(* Logix 5000 project; controller R400_500_XLS vendor 1 type 14 code 216 rev 31.11; software revision 31.01; part 28 of 32 *)
(* tags used below, declared in another part *)
   Abort1 : DINT;   // Not Used
   Ashutdown : SINT;   // Not Used
   CycExcBuffer : UDT_CYCLE;
   CycleSequence : UDT_CYCLE_SEQUENCE;
   CycleTime : DINT[11];   // Last cycle time saved in seconds
   DrnSmp : DINT;
   DRYING : DINT;   // Drying id number
   FC05_ONS : DINT;
   FINALRINSE_1 : DINT;   // Final rinse 1 id number
   FINALRINSE_9 : DINT;   // Final rinse 9 id number
   iDecimalSeparatorIndex : INT;
   M : DINT[5];   // Memory Bits
   New_Value : SINT;
   ONS_FC05 : DINT;
   ONS_FC64 : DINT;
   Print_Data : BOOL;   // Print Treatment data
   print_Door_opened_template : STRING;   // Template for the door opened message
   print_Header_template : STRING[6];   // Template for the cycle header
   Print_Speed_Water : BOOL;
   Print_TreatEnd_Start_Data : BOOL;   // 2nd treatment of the cycle is started, pirnt Treatment Completed and Treatment data
   Print_TreatStart_Data : BOOL;   // Cycle is started Print start time and treatment data of the first treatment of the cycle
   PrintBufferInjectionRate : REAL;
   printTreatString : STRING[85];   // Treatment String
   PWR_PrintBuffer : UDT_WASH;
   rBuffer : REAL[4];
   rIn_WSH61 : REAL;
   Run : DINT;
   sCRLF : STRING;
   sDecimalSeparator : STRING;
   sFll_Zero : STRING[20];
   sOut_WSH61 : STRING;
   sPrntArray : STRING[300];   // Printer String Array
   SRE3_Serial_Number : STRING;   // Serial number
   String : STRING[50];   // String
   String_Temp : STRING;
   Tmr : TIMER[107];
   Trt_PrWsh : DINT;
   WASH_1 : DINT;   // Wash 1 id number
   WASH_5 : DINT;   // Wash 5 id number
   WSH36_SecondsRemaining : DINT;
   WSH36_TotalMinutesRemaining : DINT;
   WSH36_TotalSecondsRemaining : DINT;
   WSH41_Door_opened : STRING;
   WSH41_End_signal : BOOL;   // End of cycle signal
   WSH41_Header : STRING[6];   // The header being transferred to the print queue.
   WSH41_Hour : DINT;
   WSH41_Minute : DINT;
   WSH41_ONS : SINT;
   WSH41_Second : DINT;
   WSH41_Start_signal : BOOL;   // Start cycle signal One shot rising edge
   WSH41_Temp_time : STRING[3];
   WSH41_Time_template : STRING;
   WSH41_Total_minute : DINT;
   WSH41_Total_second : DINT;
   WSH41_Total_time : STRING;
   WSH41_Zero : STRING;
   ChemConcUnit : BOOL;   // 0 = mL/L; 1 = oz/gal
   ChemicalName : STRING[9];   // Used by HMI
   CurrentUser : STRING;   // Current User
   CycleName : STRING[12];
   CyclePtr : DINT;   // Cycle Pointeur
   ENABLE : BOOL;   // Enable bit
   I_Ld_Dr_Cls_Sw : BOOL;   // Load door close
   I_Unld_Dr_Cls_Sw : BOOL;   // Unload door close
   MaintainOpenLd : BOOL;
   MaintainOpenUnld : BOOL;
   PrintIndex : DINT;
   RcvryWtrTemp : DINT;
   sCycleCounter : STRING;
   sDate : STRING;   // String current date
   sTime : STRING;   // String current time
   SumpTemp : REAL;   // Sump temperature in °C
   TempUnit : BOOL;   // Temperature Units 0= Celcius 1 = Farhenheit
   Unit : Hrdwre;   // Unit Configuration
   UnLoad : Doors;
(* MainProgram, continued *)

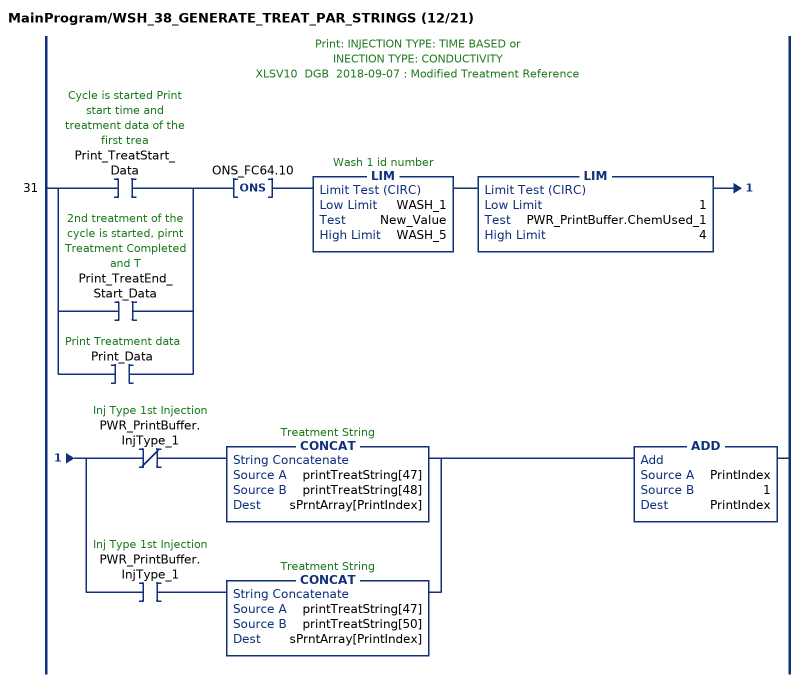
   [picture p570: MainProgram/WSH_38_GENERATE_TREAT_PAR_STRINGS rungs 31-31]
   // Print: INJECTION TYPE: TIME BASED or
   // INECTION TYPE: CONDUCTIVITY
   // XLSV10  DGB  2018-09-07 : Modified Treatment Reference
   31: [XIC(Print_TreatStart_Data) ,XIC(Print_TreatEnd_Start_Data) ,XIC(Print_Data) ]ONS(ONS_FC64.10)LIM(WASH_1,New_Value,WASH_5)LIM(1,PWR_PrintBuffer.ChemUsed_1,4)[XIO(PWR_PrintBuffer.InjType_1) CONCAT(printTreatString[47],printTreatString[48],sPrntArray[PrintIndex]) ,XIC(PWR_PrintBuffer.InjType_1) CONCAT(printTreatString[47],printTreatString[50],sPrntArray[PrintIndex]) ]ADD(PrintIndex,1,PrintIndex);
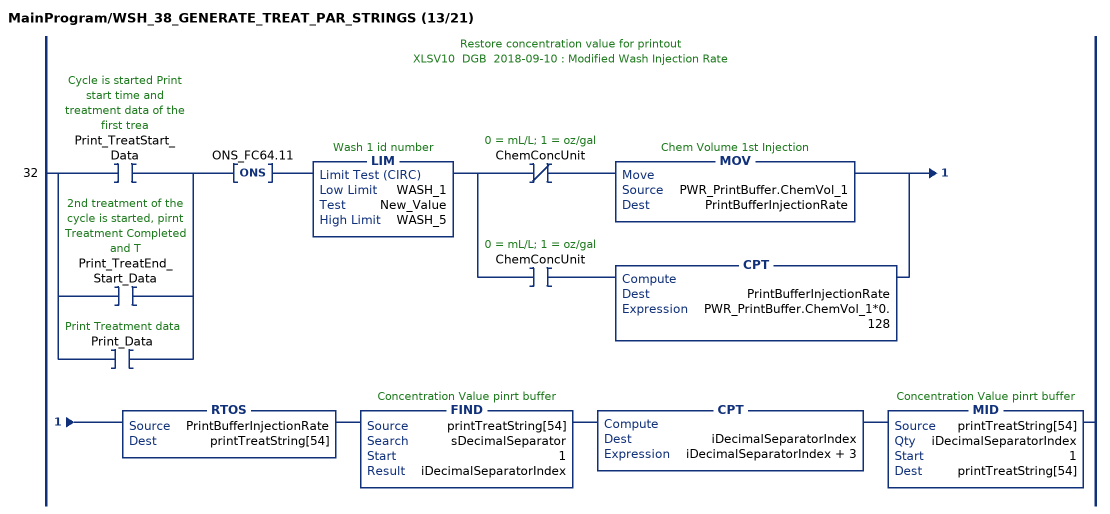
   // Restore concentration value for printout
   // XLSV10  DGB  2018-09-10 : Modified Wash Injection Rate
   32: [XIC(Print_TreatStart_Data) ,XIC(Print_TreatEnd_Start_Data) ,XIC(Print_Data) ]ONS(ONS_FC64.11)LIM(WASH_1,New_Value,WASH_5)[XIO(ChemConcUnit) MOV(PWR_PrintBuffer.ChemVol_1,PrintBufferInjectionRate) ,XIC(ChemConcUnit) CPT(PrintBufferInjectionRate,PWR_PrintBuffer.ChemVol_1*0.128) ]RTOS(PrintBufferInjectionRate,printTreatString[54])FIND(printTreatString[54],sDecimalSeparator,1,iDecimalSeparatorIndex)CPT(iDecimalSeparatorIndex,iDecimalSeparatorIndex + 3)MID(printTreatString[54],iDecimalSeparatorIndex,1,printTreatString[54]);
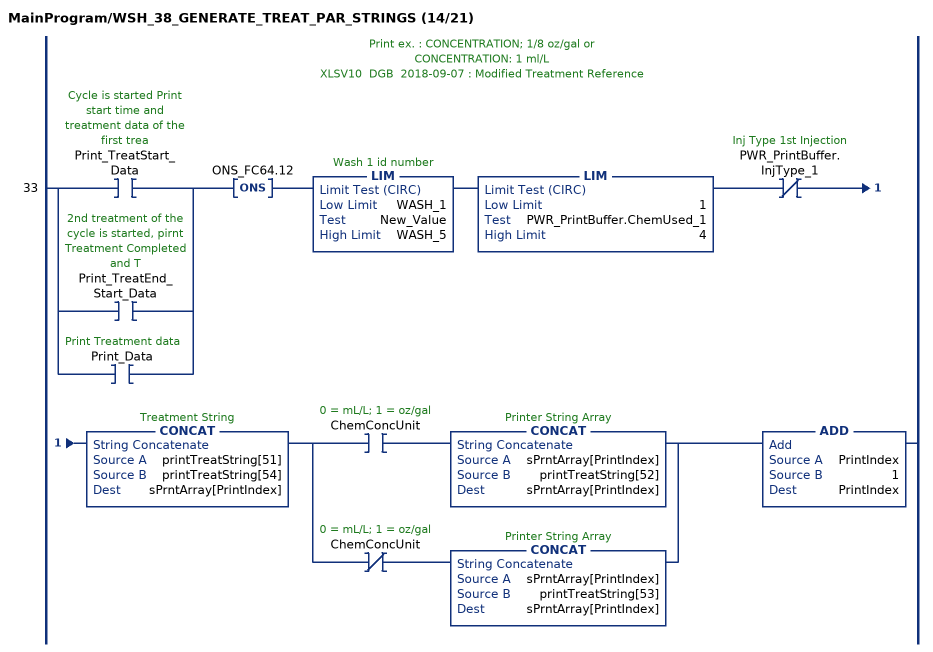
   // Print ex. : CONCENTRATION; 1/8 oz/gal or
   //         CONCENTRATION: 1 ml/L
   // XLSV10  DGB  2018-09-07 : Modified Treatment Reference
   33: [XIC(Print_TreatStart_Data) ,XIC(Print_TreatEnd_Start_Data) ,XIC(Print_Data) ]ONS(ONS_FC64.12)LIM(WASH_1,New_Value,WASH_5)LIM(1,PWR_PrintBuffer.ChemUsed_1,4)XIO(PWR_PrintBuffer.InjType_1)CONCAT(printTreatString[51],printTreatString[54],sPrntArray[PrintIndex])[XIC(ChemConcUnit) CONCAT(sPrntArray[PrintIndex],printTreatString[52],sPrntArray[PrintIndex]) ,XIO(ChemConcUnit) CONCAT(sPrntArray[PrintIndex],printTreatString[53],sPrntArray[PrintIndex]) ]ADD(PrintIndex,1,PrintIndex);
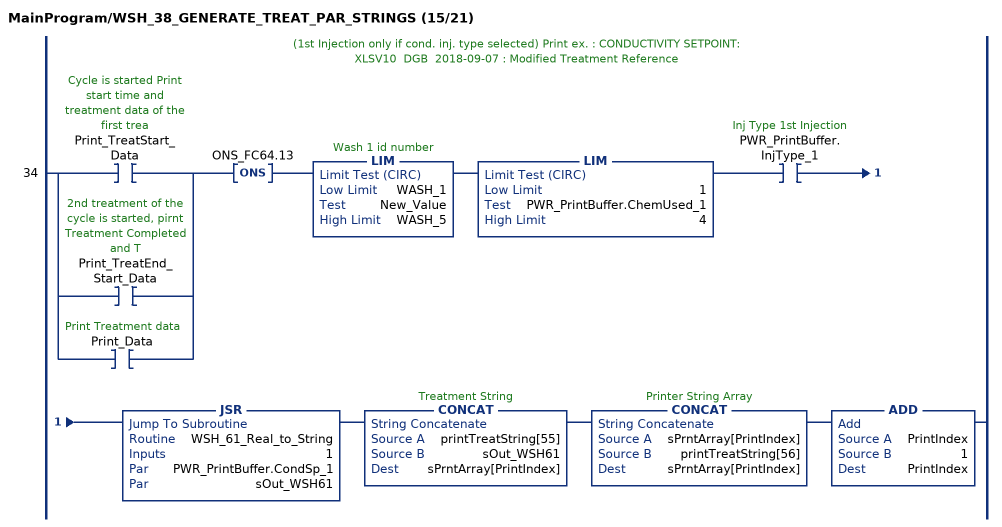
   // (1st Injection only if cond. inj. type selected) Print ex. : CONDUCTIVITY SETPOINT:
   // XLSV10  DGB  2018-09-07 : Modified Treatment Reference
   34: [XIC(Print_TreatStart_Data) ,XIC(Print_TreatEnd_Start_Data) ,XIC(Print_Data) ]ONS(ONS_FC64.13)LIM(WASH_1,New_Value,WASH_5)LIM(1,PWR_PrintBuffer.ChemUsed_1,4)XIC(PWR_PrintBuffer.InjType_1)JSR(WSH_61_Real_to_String,1,PWR_PrintBuffer.CondSp_1,sOut_WSH61)CONCAT(printTreatString[55],sOut_WSH61,sPrntArray[PrintIndex])CONCAT(sPrntArray[PrintIndex],printTreatString[56],sPrntArray[PrintIndex])ADD(PrintIndex,1,PrintIndex);
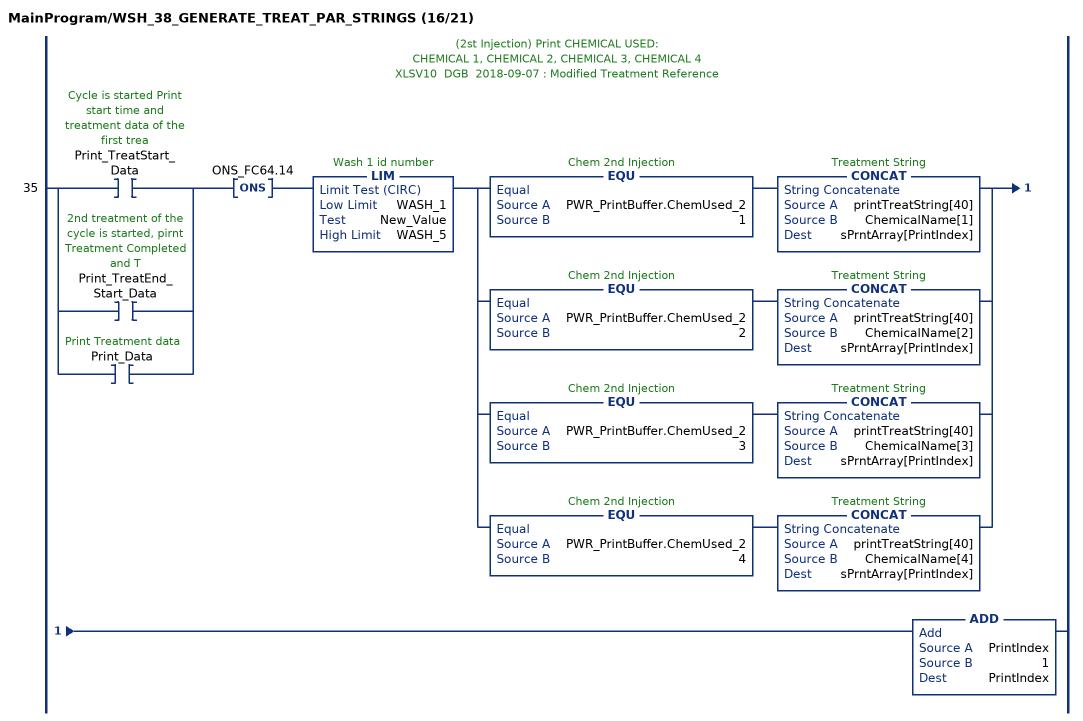
   // (2st Injection) Print CHEMICAL USED:
   //  CHEMICAL 1, CHEMICAL 2, CHEMICAL 3, CHEMICAL 4
   // XLSV10  DGB  2018-09-07 : Modified Treatment Reference
   35: [XIC(Print_TreatStart_Data) ,XIC(Print_TreatEnd_Start_Data) ,XIC(Print_Data) ]ONS(ONS_FC64.14)LIM(WASH_1,New_Value,WASH_5)[EQU(PWR_PrintBuffer.ChemUsed_2,1) CONCAT(printTreatString[40],ChemicalName[1],sPrntArray[PrintIndex]) ,EQU(PWR_PrintBuffer.ChemUsed_2,2) CONCAT(printTreatString[40],ChemicalName[2],sPrntArray[PrintIndex]) ,EQU(PWR_PrintBuffer.ChemUsed_2,3) CONCAT(printTreatString[40],ChemicalName[3],sPrntArray[PrintIndex]) ,EQU(PWR_PrintBuffer.ChemUsed_2,4) CONCAT(printTreatString[40],ChemicalName[4],sPrntArray[PrintIndex]) ]ADD(PrintIndex,1,PrintIndex);
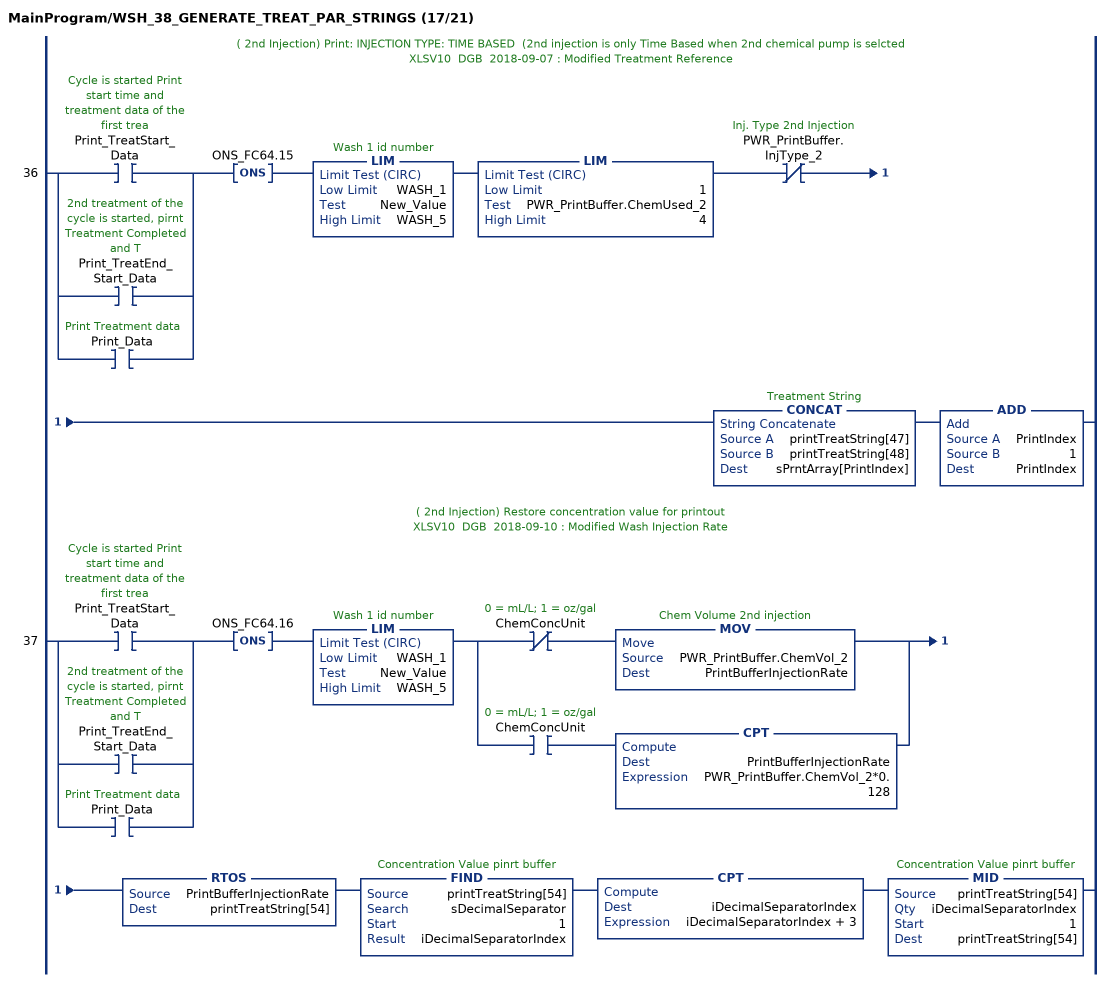
   // ( 2nd Injection) Print: INJECTION TYPE: TIME BASED  (2nd injection is only Time Based when 2nd chemical pump is selcted
   // XLSV10  DGB  2018-09-07 : Modified Treatment Reference
   36: [XIC(Print_TreatStart_Data) ,XIC(Print_TreatEnd_Start_Data) ,XIC(Print_Data) ]ONS(ONS_FC64.15)LIM(WASH_1,New_Value,WASH_5)LIM(1,PWR_PrintBuffer.ChemUsed_2,4)XIO(PWR_PrintBuffer.InjType_2)CONCAT(printTreatString[47],printTreatString[48],sPrntArray[PrintIndex])ADD(PrintIndex,1,PrintIndex);
   // ( 2nd Injection) Restore concentration value for printout
   // XLSV10  DGB  2018-09-10 : Modified Wash Injection Rate
   37: [XIC(Print_TreatStart_Data) ,XIC(Print_TreatEnd_Start_Data) ,XIC(Print_Data) ]ONS(ONS_FC64.16)LIM(WASH_1,New_Value,WASH_5)[XIO(ChemConcUnit) MOV(PWR_PrintBuffer.ChemVol_2,PrintBufferInjectionRate) ,XIC(ChemConcUnit) CPT(PrintBufferInjectionRate,PWR_PrintBuffer.ChemVol_2*0.128) ]RTOS(PrintBufferInjectionRate,printTreatString[54])FIND(printTreatString[54],sDecimalSeparator,1,iDecimalSeparatorIndex)CPT(iDecimalSeparatorIndex,iDecimalSeparatorIndex + 3)MID(printTreatString[54],iDecimalSeparatorIndex,1,printTreatString[54]);
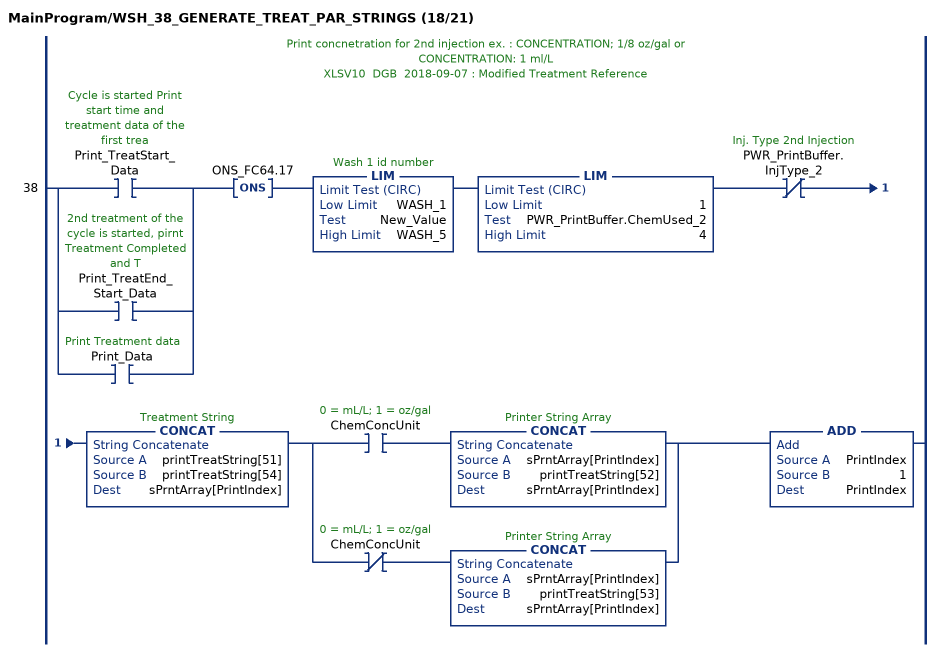
   // Print concnetration for 2nd injection ex. : CONCENTRATION; 1/8 oz/gal or
   //         CONCENTRATION: 1 ml/L
   // XLSV10  DGB  2018-09-07 : Modified Treatment Reference
   38: [XIC(Print_TreatStart_Data) ,XIC(Print_TreatEnd_Start_Data) ,XIC(Print_Data) ]ONS(ONS_FC64.17)LIM(WASH_1,New_Value,WASH_5)LIM(1,PWR_PrintBuffer.ChemUsed_2,4)XIO(PWR_PrintBuffer.InjType_2)CONCAT(printTreatString[51],printTreatString[54],sPrntArray[PrintIndex])[XIC(ChemConcUnit) CONCAT(sPrntArray[PrintIndex],printTreatString[52],sPrntArray[PrintIndex]) ,XIO(ChemConcUnit) CONCAT(sPrntArray[PrintIndex],printTreatString[53],sPrntArray[PrintIndex]) ]ADD(PrintIndex,1,PrintIndex);
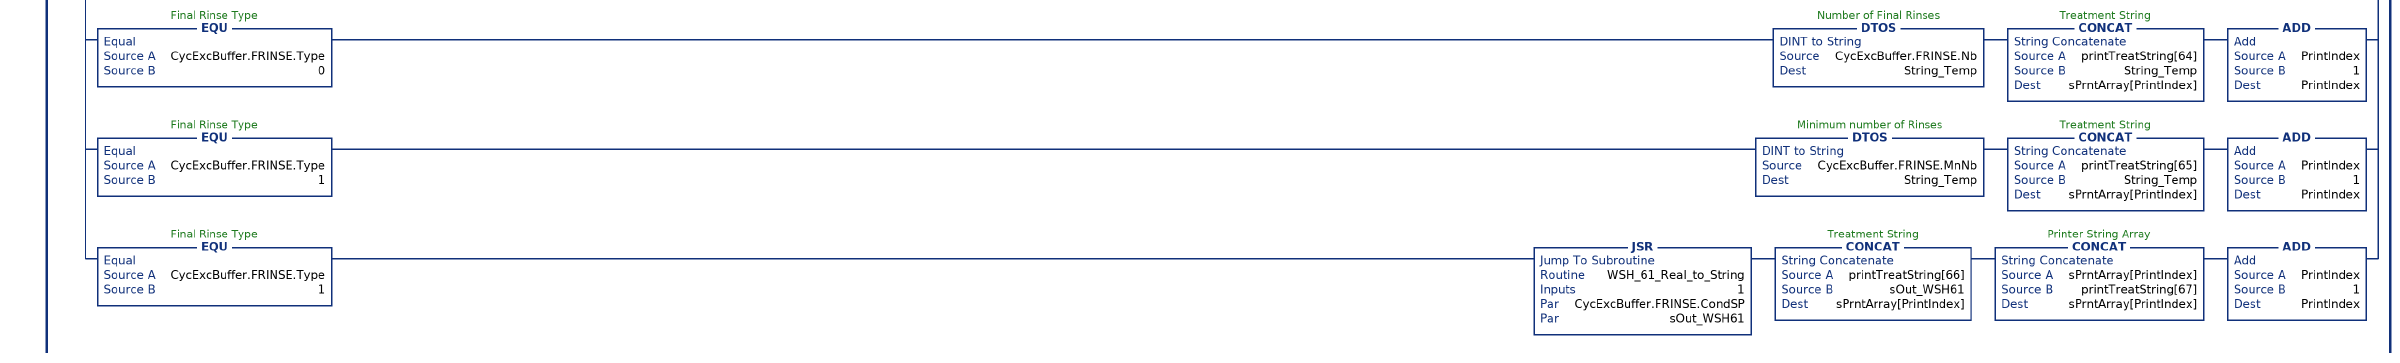
   // Print Final Rinse Data
   // XLSV10  DGB  2018-09-07 : Modified Treatment Reference
   39: [XIC(Print_TreatStart_Data) ,XIC(Print_TreatEnd_Start_Data) ,XIC(Print_Data) ]ONS(ONS_FC64.18)LIM(FINALRINSE_1,New_Value,FINALRINSE_9)[CONCAT(printTreatString[31],printTreatString[34],sPrntArray[PrintIndex]) ADD(PrintIndex,1,PrintIndex) ,XIO(CycExcBuffer.FRINSE.Heat) CONCAT(printTreatString[35],printTreatString[36],sPrntArray[PrintIndex]) ADD(PrintIndex,1,PrintIndex) ,XIC(CycExcBuffer.FRINSE.Heat) XIO(TempUnit) MOV(CycExcBuffer.FRINSE.Tmp,rIn_WSH61) JSR(WSH_61_Real_to_String,1,rIn_WSH61,sOut_WSH61) CONCAT(printTreatString[35],sOut_WSH61,sPrntArray[PrintIndex]) CONCAT(sPrntArray[PrintIndex],printTreatString[37],sPrntArray[PrintIndex]) ADD(PrintIndex,1,PrintIndex) ,XIC(CycExcBuffer.FRINSE.Heat) XIC(TempUnit) MOV(CycExcBuffer.FRINSE.Tmp,rBuffer[3]) CPT(rIn_WSH61,rBuffer[3]*1.8+32) JSR(WSH_61_Real_to_String,1,rIn_WSH61,sOut_WSH61) CONCAT(printTreatString[35],sOut_WSH61,sPrntArray[PrintIndex]) CONCAT(sPrntArray[PrintIndex],printTreatString[38],sPrntArray[PrintIndex]) ADD(PrintIndex,1,PrintIndex) ,XIO(CycExcBuffer.FRINSE.Drn) CONCAT(printTreatString[57],printTreatString[59],sPrntArray[PrintIndex]) ADD(PrintIndex,1,PrintIndex) ,XIC(CycExcBuffer.FRINSE.Drn) CONCAT(printTreatString[57],printTreatString[58],sPrntArray[PrintIndex]) ADD(PrintIndex,1,PrintIndex) ,XIC(CycExcBuffer.FRINSE.Recirc) CONCAT(printTreatString[60],printTreatString[58],sPrntArray[PrintIndex]) ADD(PrintIndex,1,PrintIndex) ,XIO(CycExcBuffer.FRINSE.Recirc) CONCAT(printTreatString[60],printTreatString[59],sPrntArray[PrintIndex]) ADD(PrintIndex,1,PrintIndex) ,[LEQ(CycExcBuffer.FRINSE.Tmin,9) DTOS(CycExcBuffer.FRINSE.Tmin,String_Temp) CONCAT(sFll_Zero[0],String_Temp,String_Temp) ,GRT(CycExcBuffer.FRINSE.Tmin,9) DTOS(CycExcBuffer.FRINSE.Tmin,String_Temp) ] CONCAT(printTreatString[39],String_Temp,sPrntArray[PrintIndex]) CONCAT(sPrntArray[PrintIndex],String[14],sPrntArray[PrintIndex]) [LEQ(CycExcBuffer.FRINSE.Tsec,9) DTOS(CycExcBuffer.FRINSE.Tsec,String_Temp) CONCAT(sFll_Zero[0],String_Temp,String_Temp) ,GRT(CycExcBuffer.FRINSE.Tsec,9) DTOS(CycExcBuffer.FRINSE.Tsec,String_Temp) ] CONCAT(sPrntArray[PrintIndex],String_Temp,sPrntArray[PrintIndex]) ADD(PrintIndex,1,PrintIndex) ,EQU(CycExcBuffer.FRINSE.Type,0) CONCAT(printTreatString[61],printTreatString[62],sPrntArray[PrintIndex]) ADD(PrintIndex,1,PrintIndex) ,EQU(CycExcBuffer.FRINSE.Type,1) CONCAT(printTreatString[61],printTreatString[63],sPrntArray[PrintIndex]) ADD(PrintIndex,1,PrintIndex) ,EQU(CycExcBuffer.FRINSE.Type,0) DTOS(CycExcBuffer.FRINSE.Nb,String_Temp) CONCAT(printTreatString[64],String_Temp,sPrntArray[PrintIndex]) ADD(PrintIndex,1,PrintIndex) ,EQU(CycExcBuffer.FRINSE.Type,1) DTOS(CycExcBuffer.FRINSE.MnNb,String_Temp) CONCAT(printTreatString[65],String_Temp,sPrntArray[PrintIndex]) ADD(PrintIndex,1,PrintIndex) ,EQU(CycExcBuffer.FRINSE.Type,1) JSR(WSH_61_Real_to_String,1,CycExcBuffer.FRINSE.CondSP,sOut_WSH61) CONCAT(printTreatString[66],sOut_WSH61,sPrntArray[PrintIndex]) CONCAT(sPrntArray[PrintIndex],printTreatString[67],sPrntArray[PrintIndex]) ADD(PrintIndex,1,PrintIndex) ];
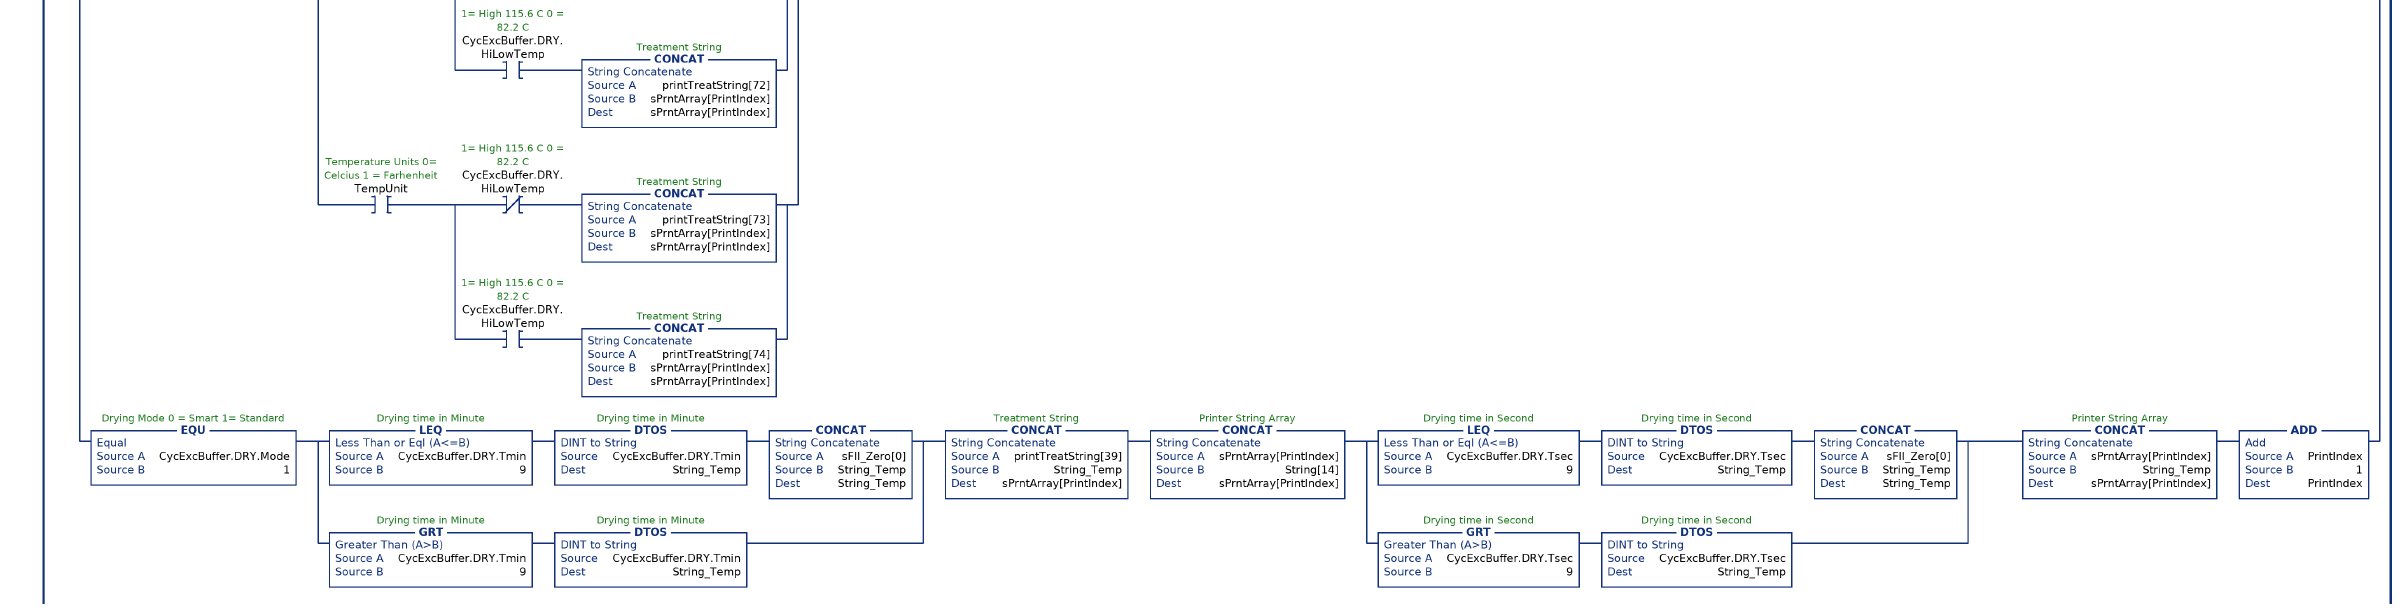
   // Print Drying Data
   // XLSV10  DGB  2018-09-07 : Modified Treatment Reference  and Changed Regular Low Temperature
   40: [XIC(Print_TreatStart_Data) ,XIC(Print_TreatEnd_Start_Data) ,XIC(Print_Data) ]ONS(ONS_FC64.19)EQU(New_Value,DRYING)[EQU(CycExcBuffer.DRY.Mode,0) CONCAT(printTreatString[68],printTreatString[69],sPrntArray[PrintIndex]) ADD(PrintIndex,1,PrintIndex) ,EQU(CycExcBuffer.DRY.Mode,1) CONCAT(printTreatString[68],printTreatString[70],sPrntArray[PrintIndex]) ADD(PrintIndex,1,PrintIndex) ,EQU(CycExcBuffer.DRY.Mode,0) XIO(CycExcBuffer.DRY.HeatSensitive) CONCAT(printTreatString[28],printTreatString[29],sPrntArray[PrintIndex]) ADD(PrintIndex,1,PrintIndex) ,EQU(CycExcBuffer.DRY.Mode,0) XIC(CycExcBuffer.DRY.HeatSensitive) CONCAT(printTreatString[28],printTreatString[75],sPrntArray[PrintIndex]) ADD(PrintIndex,1,PrintIndex) ,EQU(CycExcBuffer.DRY.Mode,1) [XIO(TempUnit) [XIO(CycExcBuffer.DRY.HiLowTemp) CONCAT(printTreatString[71],sPrntArray[PrintIndex],sPrntArray[PrintIndex]) ,XIC(CycExcBuffer.DRY.HiLowTemp) CONCAT(printTreatString[72],sPrntArray[PrintIndex],sPrntArray[PrintIndex]) ] ,XIC(TempUnit) [XIO(CycExcBuffer.DRY.HiLowTemp) CONCAT(printTreatString[73],sPrntArray[PrintIndex],sPrntArray[PrintIndex]) ,XIC(CycExcBuffer.DRY.HiLowTemp) CONCAT(printTreatString[74],sPrntArray[PrintIndex],sPrntArray[PrintIndex]) ] ] ADD(PrintIndex,1,PrintIndex) ,EQU(CycExcBuffer.DRY.Mode,1) [LEQ(CycExcBuffer.DRY.Tmin,9) DTOS(CycExcBuffer.DRY.Tmin,String_Temp) CONCAT(sFll_Zero[0],String_Temp,String_Temp) ,GRT(CycExcBuffer.DRY.Tmin,9) DTOS(CycExcBuffer.DRY.Tmin,String_Temp) ] CONCAT(printTreatString[39],String_Temp,sPrntArray[PrintIndex]) CONCAT(sPrntArray[PrintIndex],String[14],sPrntArray[PrintIndex]) [LEQ(CycExcBuffer.DRY.Tsec,9) DTOS(CycExcBuffer.DRY.Tsec,String_Temp) CONCAT(sFll_Zero[0],String_Temp,String_Temp) ,GRT(CycExcBuffer.DRY.Tsec,9) DTOS(CycExcBuffer.DRY.Tsec,String_Temp) ] CONCAT(sPrntArray[PrintIndex],String_Temp,sPrntArray[PrintIndex]) ADD(PrintIndex,1,PrintIndex) ];
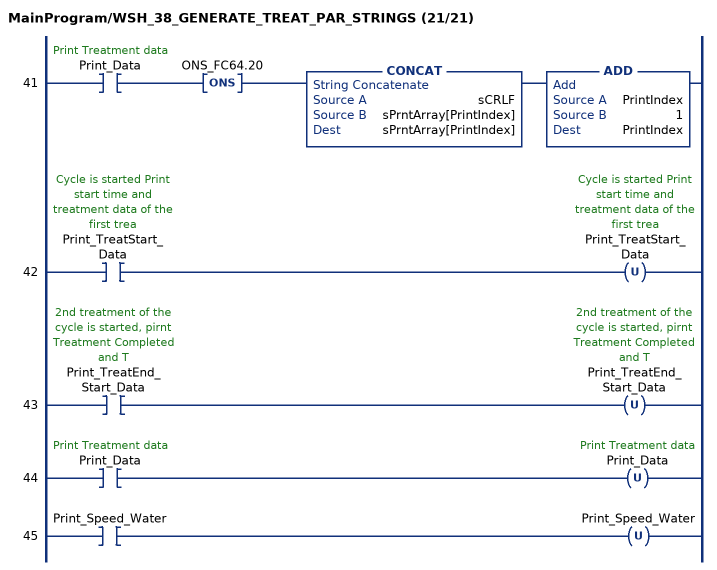
   41: XIC(Print_Data)ONS(ONS_FC64.20)CONCAT(sCRLF,sPrntArray[PrintIndex],sPrntArray[PrintIndex])ADD(PrintIndex,1,PrintIndex);
   42: XIC(Print_TreatStart_Data)OTU(Print_TreatStart_Data);
   43: XIC(Print_TreatEnd_Start_Data)OTU(Print_TreatEnd_Start_Data);
   44: XIC(Print_Data)OTU(Print_Data);
   45: XIC(Print_Speed_Water)OTU(Print_Speed_Water);
END_ROUTINE

ROUTINE WSH_41_Generate_cycle_header_footer   (* ladder *)
// This routine generates the cycle header and footer
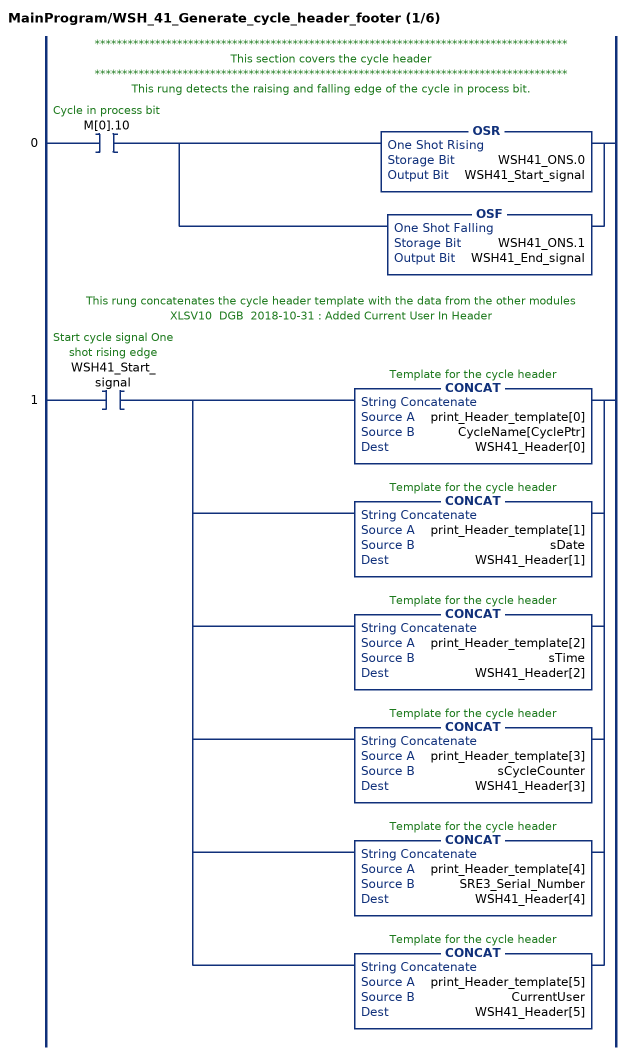
   // **************************************************************************************
   // This section covers the cycle header
   // **************************************************************************************
   // This rung detects the raising and falling edge of the cycle in process bit.
   0: XIC(M[0].10)[OSR(WSH41_ONS.0,WSH41_Start_signal) ,OSF(WSH41_ONS.1,WSH41_End_signal) ];
   // This rung concatenates the cycle header template with the data from the other modules
   // XLSV10  DGB  2018-10-31 : Added Current User In Header
   1: XIC(WSH41_Start_signal)[CONCAT(print_Header_template[0],CycleName[CyclePtr],WSH41_Header[0]) ,CONCAT(print_Header_template[1],sDate,WSH41_Header[1]) ,CONCAT(print_Header_template[2],sTime,WSH41_Header[2]) ,CONCAT(print_Header_template[3],sCycleCounter,WSH41_Header[3]) ,CONCAT(print_Header_template[4],SRE3_Serial_Number,WSH41_Header[4]) ,CONCAT(print_Header_template[5],CurrentUser,WSH41_Header[5]) ];
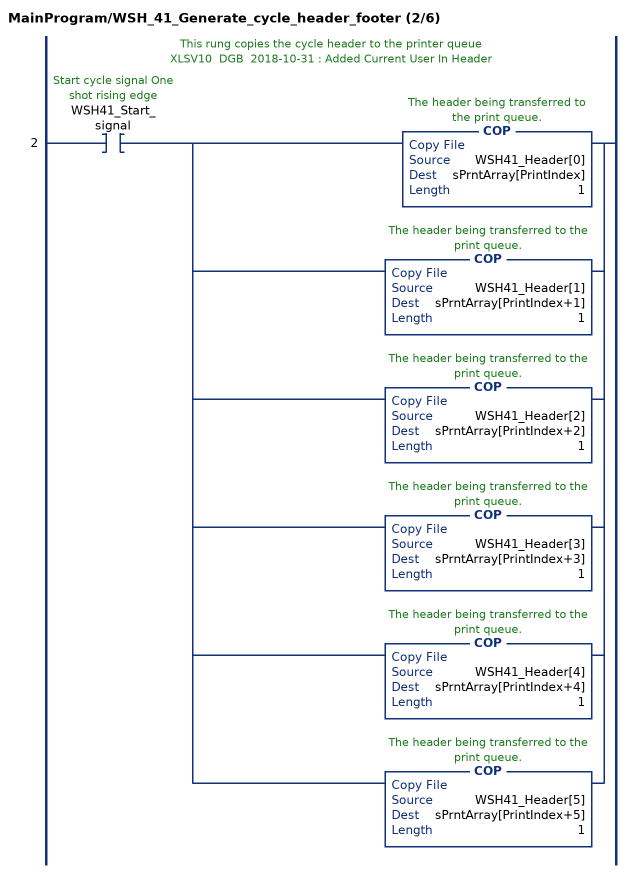
   // This rung copies the cycle header to the printer queue
   // XLSV10  DGB  2018-10-31 : Added Current User In Header
   2: XIC(WSH41_Start_signal)[COP(WSH41_Header[0],sPrntArray[PrintIndex],1) ,COP(WSH41_Header[1],sPrntArray[PrintIndex+1],1) ,COP(WSH41_Header[2],sPrntArray[PrintIndex+2],1) ,COP(WSH41_Header[3],sPrntArray[PrintIndex+3],1) ,COP(WSH41_Header[4],sPrntArray[PrintIndex+4],1) ,COP(WSH41_Header[5],sPrntArray[PrintIndex+5],1) ];
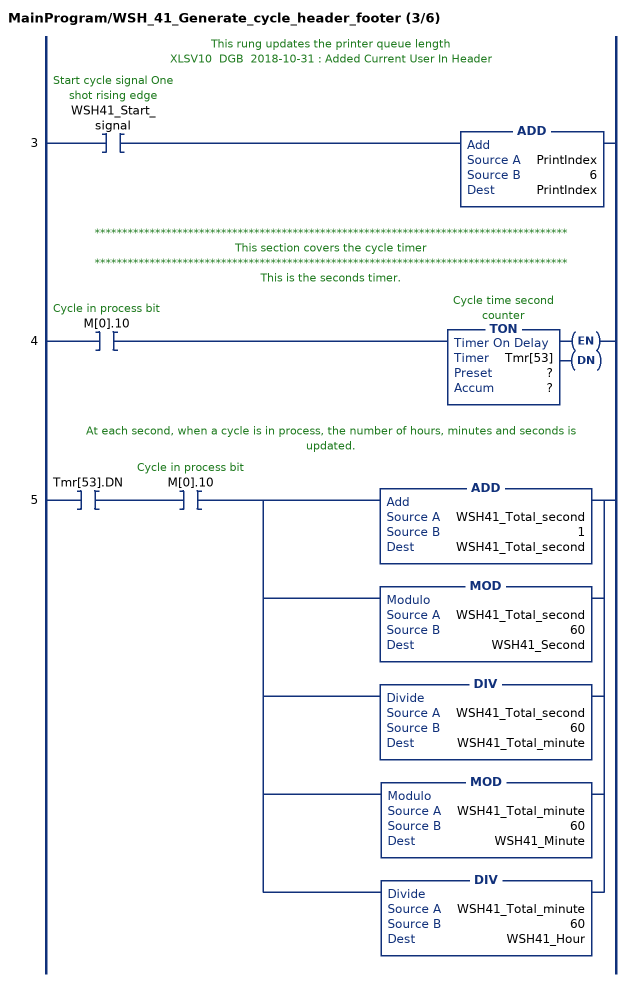
   // This rung updates the printer queue length
   // XLSV10  DGB  2018-10-31 : Added Current User In Header
   3: XIC(WSH41_Start_signal)ADD(PrintIndex,6,PrintIndex);
   // **************************************************************************************
   // This section covers the cycle timer
   // **************************************************************************************
   // This is the seconds timer.
   4: XIC(M[0].10)TON(Tmr[53],?,?);
   // At each second, when a cycle is in process, the number of hours, minutes and seconds is updated.
   5: XIC(Tmr[53].DN)XIC(M[0].10)[ADD(WSH41_Total_second,1,WSH41_Total_second) ,MOD(WSH41_Total_second,60,WSH41_Second) ,DIV(WSH41_Total_second,60,WSH41_Total_minute) ,MOD(WSH41_Total_minute,60,WSH41_Minute) ,DIV(WSH41_Total_minute,60,WSH41_Hour) ];
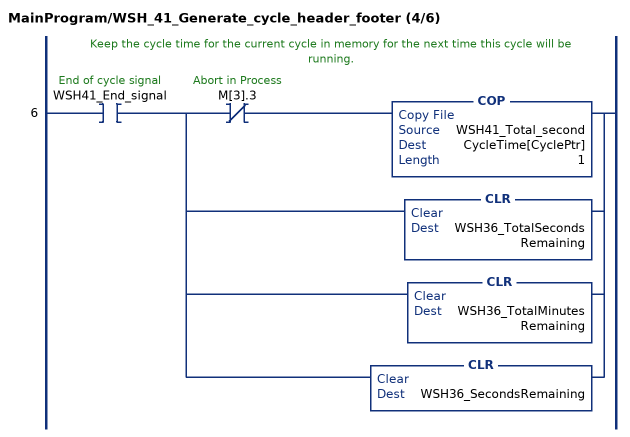
   // Keep the cycle time for the current cycle in memory for the next time this cycle will be running.
   6: XIC(WSH41_End_signal)[XIO(M[3].3) COP(WSH41_Total_second,CycleTime[CyclePtr],1) ,CLR(WSH36_TotalSecondsRemaining) ,CLR(WSH36_TotalMinutesRemaining) ,CLR(WSH36_SecondsRemaining) ];
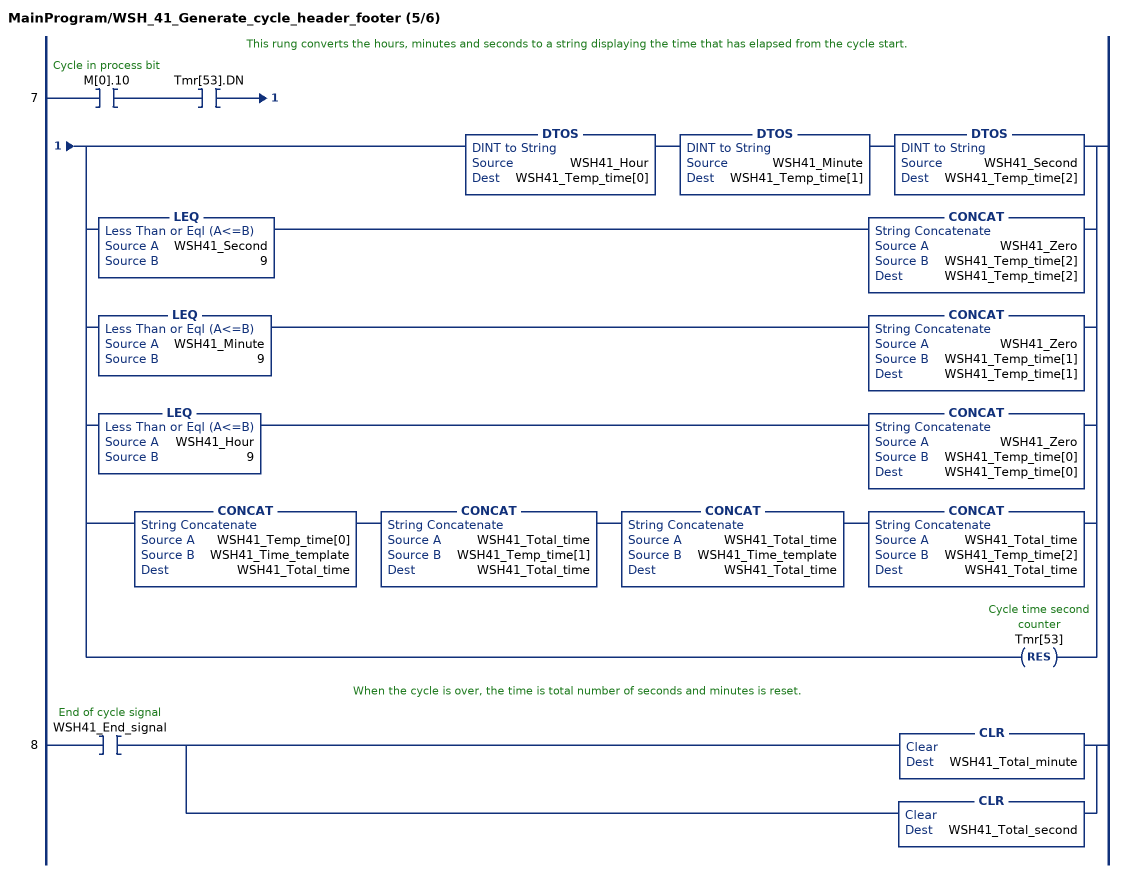
   // This rung converts the hours, minutes and seconds to a string displaying the time that has elapsed from the cycle start.
   7: XIC(M[0].10)XIC(Tmr[53].DN)[DTOS(WSH41_Hour,WSH41_Temp_time[0]) DTOS(WSH41_Minute,WSH41_Temp_time[1]) DTOS(WSH41_Second,WSH41_Temp_time[2]) ,LEQ(WSH41_Second,9) CONCAT(WSH41_Zero,WSH41_Temp_time[2],WSH41_Temp_time[2]) ,LEQ(WSH41_Minute,9) CONCAT(WSH41_Zero,WSH41_Temp_time[1],WSH41_Temp_time[1]) ,LEQ(WSH41_Hour,9) CONCAT(WSH41_Zero,WSH41_Temp_time[0],WSH41_Temp_time[0]) ,CONCAT(WSH41_Temp_time[0],WSH41_Time_template,WSH41_Total_time) CONCAT(WSH41_Total_time,WSH41_Temp_time[1],WSH41_Total_time) CONCAT(WSH41_Total_time,WSH41_Time_template,WSH41_Total_time) CONCAT(WSH41_Total_time,WSH41_Temp_time[2],WSH41_Total_time) ,RES(Tmr[53]) ];
   // When the cycle is over, the time is total number of seconds and minutes is reset.
   8: XIC(WSH41_End_signal)[CLR(WSH41_Total_minute) ,CLR(WSH41_Total_second) ];
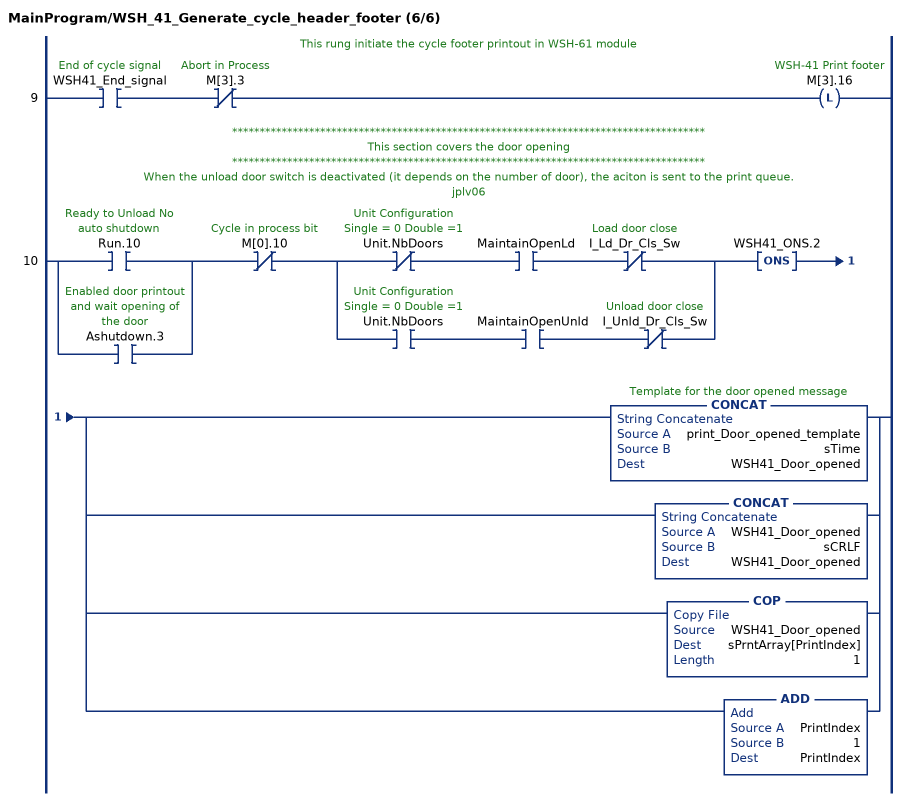
   // This rung initiate the cycle footer printout in WSH-61 module
   9: XIC(WSH41_End_signal)XIO(M[3].3)OTL(M[3].16);
   // **************************************************************************************
   // This section covers the door opening
   // **************************************************************************************
   // When the unload door switch is deactivated (it depends on the number of door), the aciton is sent to the print queue.
   // jplv06
   10: [XIC(Run.10) ,XIC(Ashutdown.3) ]XIO(M[0].10)[XIO(Unit.NbDoors) XIC(MaintainOpenLd) XIO(I_Ld_Dr_Cls_Sw) ,XIC(Unit.NbDoors) XIC(MaintainOpenUnld) XIO(I_Unld_Dr_Cls_Sw) ]ONS(WSH41_ONS.2)[CONCAT(print_Door_opened_template,sTime,WSH41_Door_opened) ,CONCAT(WSH41_Door_opened,sCRLF,WSH41_Door_opened) ,COP(WSH41_Door_opened,sPrntArray[PrintIndex],1) ,ADD(PrintIndex,1,PrintIndex) ];
END_ROUTINE

ROUTINE WSH_55_TRT_PW   (* ladder *)
// This module call routine to perform
// Pre-Wah treatments
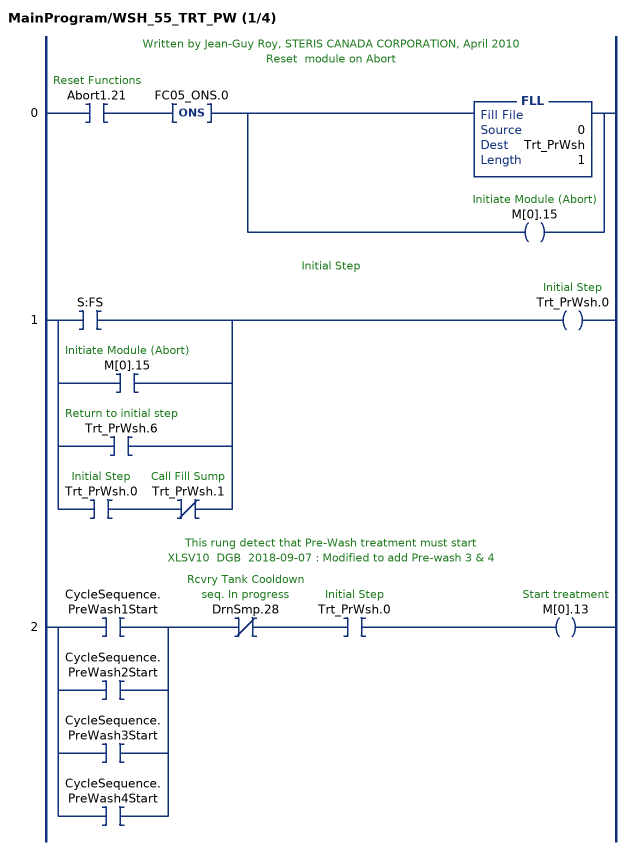
   // Written by Jean-Guy Roy, STERIS CANADA CORPORATION, April 2010
   // Reset  module on Abort
   0: XIC(Abort1.21)ONS(FC05_ONS.0)[FLL(0,Trt_PrWsh,1) ,OTE(M[0].15) ];
   // Initial Step
   1: [XIC(S:FS) ,XIC(M[0].15) ,XIC(Trt_PrWsh.6) ,XIC(Trt_PrWsh.0) XIO(Trt_PrWsh.1) ]OTE(Trt_PrWsh.0);
   // This rung detect that Pre-Wash treatment must start
   // XLSV10  DGB  2018-09-07 : Modified to add Pre-wash 3 & 4
   2: [XIC(CycleSequence.PreWash1Start) ,XIC(CycleSequence.PreWash2Start) ,XIC(CycleSequence.PreWash3Start) ,XIC(CycleSequence.PreWash4Start) ]XIO(DrnSmp.28)XIC(Trt_PrWsh.0)OTE(M[0].13);
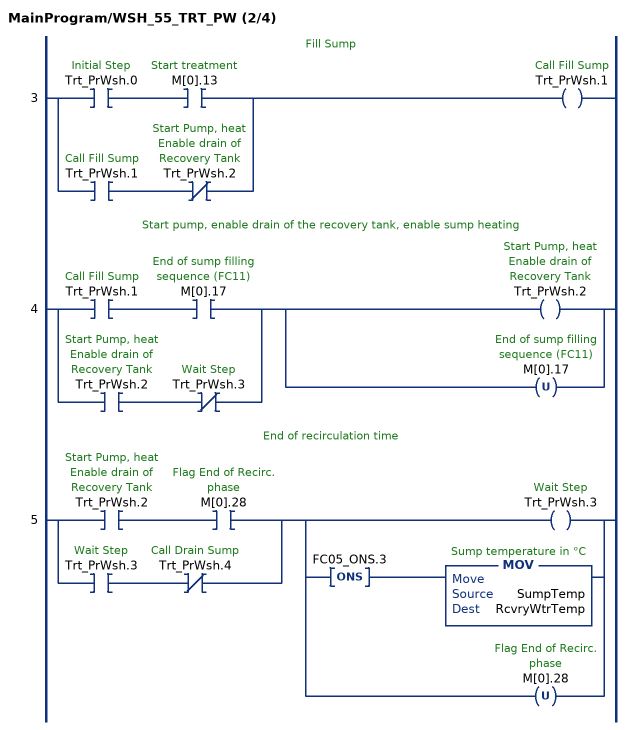
   // Fill Sump
   3: [XIC(Trt_PrWsh.0) XIC(M[0].13) ,XIC(Trt_PrWsh.1) XIO(Trt_PrWsh.2) ]OTE(Trt_PrWsh.1);
   // Start pump, enable drain of the recovery tank, enable sump heating
   4: [XIC(Trt_PrWsh.1) XIC(M[0].17) ,XIC(Trt_PrWsh.2) XIO(Trt_PrWsh.3) ][OTE(Trt_PrWsh.2) ,OTU(M[0].17) ];
   // End of recirculation time
   5: [XIC(Trt_PrWsh.2) XIC(M[0].28) ,XIC(Trt_PrWsh.3) XIO(Trt_PrWsh.4) ][OTE(Trt_PrWsh.3) ,ONS(FC05_ONS.3) MOV(SumpTemp,RcvryWtrTemp) ,OTU(M[0].28) ];
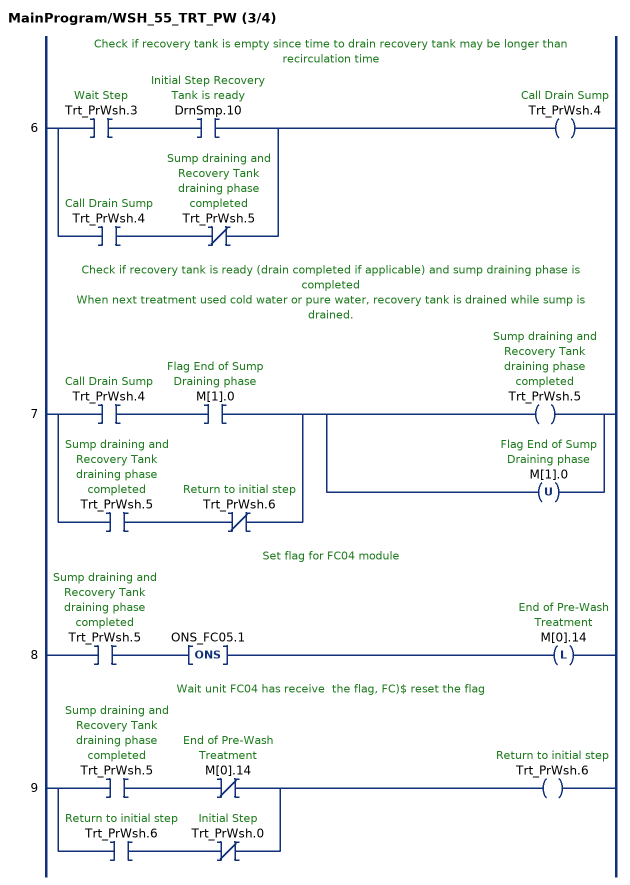
   // Check if recovery tank is empty since time to drain recovery tank may be longer than recirculation time
   6: [XIC(Trt_PrWsh.3) XIC(DrnSmp.10) ,XIC(Trt_PrWsh.4) XIO(Trt_PrWsh.5) ]OTE(Trt_PrWsh.4);
   // Check if recovery tank is ready (drain completed if applicable) and sump draining phase is completed
   // When next treatment used cold water or pure water, recovery tank is drained while sump is drained.
   7: [XIC(Trt_PrWsh.4) XIC(M[1].0) ,XIC(Trt_PrWsh.5) XIO(Trt_PrWsh.6) ][OTE(Trt_PrWsh.5) ,OTU(M[1].0) ];
   // Set flag for FC04 module
   8: XIC(Trt_PrWsh.5)ONS(ONS_FC05.1)OTL(M[0].14);
   // Wait unit FC04 has receive  the flag, FC)$ reset the flag
   9: [XIC(Trt_PrWsh.5) XIO(M[0].14) ,XIC(Trt_PrWsh.6) XIO(Trt_PrWsh.0) ]OTE(Trt_PrWsh.6);
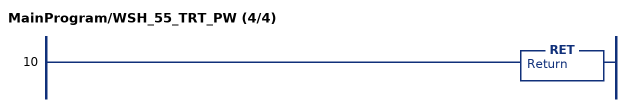
   10: RET();
END_ROUTINE
